FUNCTION_BLOCK FB_PERIPHERY_REF_1
VAR_INPUT

END_VAR
VAR_OUTPUT

END_VAR
VAR_IN_OUT

END_VAR
VAR

END_VAR

;

END_FUNCTION_BLOCK

(* stored: Version 1.1.0.1, ProductVersion 3.1.4024.15
   POU FB_PERIPHERY_REF_1: Id {dbffa441-33d1-4615-9356-5a5b76714dbd}, SpecialFunc None *)
